// TIA Portal V20 export
// export: Created 2026-10-20T12:47:33.6136507Z, ExportSetting WithDefaults, DisplayName Totally Integrated Automation Portal, DisplayVersion V20 Update 6, DisplayName TIA Portal Openness, DisplayVersion V20 Update 6, DisplayName TIA Portal Version Control Interface, DisplayVersion V20 Update 6, DisplayName SINAMICS Startdrive Advanced, DisplayVersion V20 SP1, DisplayName SINAMICS Startdrive G130, G150, S120, S150, SINAMICS MV, G220, S200, S210, DisplayVersion V20 SP1, DisplayName SINAMICS Startdrive G110M, G120, G120C, G120D, G120P, G115D, DisplayVersion V20 SP1, DisplayName STEP 7 Professional, DisplayVersion V20 Update 6, DisplayName STEP 7 Safety, DisplayVersion V20 Update 2, DisplayName WinCC Basic/Comfort/Advanced, DisplayVersion V20 Update 6, DisplayName WinCC Unified, DisplayVersion V20 Update 6
FUNCTION_BLOCK "FB_HeartBeat"   // FB25, SCL
{ S7_Optimized_Access := 'TRUE' }
VERSION : 0.1
// stored: AutoNumber true, IsIECCheckEnabled false, IsRetainMemResEnabled false, MemoryReserve 100, SetENOAutomatically false, UDAEnableTagReadback false
   VAR_INPUT
      PC_HeartBeat : Word;
   END_VAR
   VAR_OUTPUT
      PLC_HeartBeat : Word;
      PC_Disconnected : Bool;
   END_VAR
   VAR
      TimeOut : TON_TIME;
      "Timer" { S7_SetPoint := 'True'} : TON_TIME;
      PC_Heartbeat_old : Word;
      StartTimerBit : Bool := FALSE;
   END_VAR
BEGIN
   #Timer(IN := #StartTimerBit, //
          PT := t#250ms);
   IF NOT #StartTimerBit THEN
       #StartTimerBit := TRUE;
   END_IF;
   #Timer(IN := #StartTimerBit, //
          PT := t#250ms);
   IF #Timer.Q THEN
       #StartTimerBit := FALSE;
       RESET_TIMER(#Timer);
       #PLC_HeartBeat += 1;
   END_IF;
   //Time Out Timer
   #TimeOut(IN := #PC_HeartBeat = #PC_Heartbeat_old,
            PT := t#10s);
   #PC_Heartbeat_old := #PC_HeartBeat;
   #PC_Disconnected := #TimeOut.Q; // if time out set PC_Disconnected
END_FUNCTION_BLOCK
